(* IEC 61131-3 sources: plc-vscode/tests/st/all/rusty/tests/lit/multi/cross_file_hardware_alias_1307, 2 files *)

(* ---- file1.st ---- *)
VAR_GLOBAL
    foo AT %IX1.2.3.4 : BOOL;
END_VAR

FUNCTION main : DINT
    // Confirm the alias is wired by writing through `foo` and reading it back.
    // file2.st declares `bar` at the same hardware address, so the two names
    // must share the same backing storage (`__PI_1_2_3_4`).
    foo := TRUE;
    IF foo THEN
        printf('aliased$N');
    END_IF;
    main := 0;
END_FUNCTION

(* ---- file2.st ---- *)
// Declared in a separate compilation unit at the same hardware address as
// file1.st's `foo`. Without the cross-unit dedup of synthetic `__PI_*`
// globals, this used to fail to link with an ambiguous-symbol error
// (#1307).
VAR_GLOBAL
    bar AT %IX1.2.3.4 : BOOL;
END_VAR
